(* IEC 61131-3 sources: iolistgen/tests_support/pl_stub/src/DUTs/ControlValve, 5 files *)

(* ---- E_CvAlarm.dut.st ---- *)
// Назначение: заглушка plc-process-lib 1.0.0 для проверки типов сгенерированного кода без CODESYS
//             (API.md, раздел 4.1); не библиотека — тел и внутренних переменных нет
// Автор:      kr0nsch
// Версия:     1.0.0 (выпуск библиотеки)
// Документ:   docs/GENERATORS.md, раздел «Проверка ST без CODESYS»
{attribute 'qualified_only'}
TYPE E_CvAlarm :
(
    Deviation := 0,
    FbFailure := 1,
    PositionerFault := 2,
    InterlockAct := 3
) UINT;
END_TYPE

(* ---- E_CvFaultAction.dut.st ---- *)
// Назначение: заглушка plc-process-lib 1.0.0 для проверки типов сгенерированного кода без CODESYS
//             (API.md, раздел 16.1); не библиотека — тел и внутренних переменных нет
// Автор:      kr0nsch
// Версия:     1.0.0 (выпуск библиотеки)
// Документ:   docs/GENERATORS.md, раздел «Проверка ST без CODESYS»
{attribute 'qualified_only'}
{attribute 'strict'}
TYPE E_CvFaultAction :
(
    Hold := 0,
    SafePos := 1
) INT;
END_TYPE

(* ---- ST_ControlValveCfg.dut.st ---- *)
// Назначение: заглушка plc-process-lib 1.0.0 для проверки типов сгенерированного кода без CODESYS
//             (API.md, раздел 16.1); не библиотека — тел и внутренних переменных нет
// Автор:      kr0nsch
// Версия:     1.0.0 (выпуск библиотеки)
// Документ:   docs/GENERATORS.md, раздел «Проверка ST без CODESYS»
{attribute 'qualified_only'}
TYPE ST_ControlValveCfg :
STRUCT
    rOutMin_pct     : REAL := 0.0;
    rOutMax_pct     : REAL := 100.0;
    rRateUp_pctps   : REAL := 0.0;
    rRateDown_pctps : REAL := 0.0;
    rTightShut_pct  : REAL := 0.0;
    xOutInvert      : BOOL := FALSE;
    rSafePos_pct    : REAL := 0.0;
    eFaultAction    : E_CvFaultAction := E_CvFaultAction.Hold;
    xFbUsed         : BOOL := FALSE;
    rDevMax_pct     : REAL := 5.0;
    tDev            : TIME := T#30S;
    xDevIsFault     : BOOL := FALSE;
    wInterlockMask  : WORD := 16#FFFF;
    udiAlarmIdBase  : UDINT := 0;
    // lint:allow STL007 имя массива по контракту API.md (префикс a + тип элемента)
    astAlarm       : ARRAY[0..GVL_Const.DEV_ALARMS_MAX - 1] OF ST_AlarmCfg := [
            (ePriority := E_AlarmPriority.Low),
            (ePriority := E_AlarmPriority.Low),
            (ePriority := E_AlarmPriority.Medium),
            (ePriority := E_AlarmPriority.None),
            (ePriority := E_AlarmPriority.None),
            (ePriority := E_AlarmPriority.None),
            (ePriority := E_AlarmPriority.None),
            (ePriority := E_AlarmPriority.None)];
END_STRUCT
END_TYPE

(* ---- ST_ControlValveCmd.dut.st ---- *)
// Назначение: заглушка plc-process-lib 1.0.0 для проверки типов сгенерированного кода без CODESYS
//             (API.md, раздел 16.1); не библиотека — тел и внутренних переменных нет
// Автор:      kr0nsch
// Версия:     1.0.0 (выпуск библиотеки)
// Документ:   docs/GENERATORS.md, раздел «Проверка ST без CODESYS»
{attribute 'qualified_only'}
TYPE ST_ControlValveCmd :
STRUCT
    stCommon      : ST_DeviceCmd;
    rPosSpMan_pct : REAL;
END_STRUCT
END_TYPE

(* ---- ST_ControlValveSts.dut.st ---- *)
// Назначение: заглушка plc-process-lib 1.0.0 для проверки типов сгенерированного кода без CODESYS
//             (API.md, раздел 16.1); не библиотека — тел и внутренних переменных нет
// Автор:      kr0nsch
// Версия:     1.0.0 (выпуск библиотеки)
// Документ:   docs/GENERATORS.md, раздел «Проверка ST без CODESYS»
{attribute 'qualified_only'}
TYPE ST_ControlValveSts :
STRUCT
    stCommon       : ST_DeviceSts;
    rPosSp_pct     : REAL;
    rOut_pct       : REAL;
    rOut_mA        : REAL;
    rPosFb_pct     : REAL;
    rDeviation_pct : REAL;
    wInterlock     : WORD;
    uiFirstOut     : UINT;
END_STRUCT
END_TYPE
